// TIA Portal project "exografcet2" (V16)

(* hardware
DEVICE "Station S7-1200_1"  S7-1200 Station
   slot 0: "Châssis_0"  S7-1200 Rack  Rack  V1.0
   slot 1: "PLC_1"  CPU 1214C AC/DC/Rly  6ES7 214-1BG40-0XB0  V4.4
*)

// ===== PLC "PLC_1"  CPU 1214C AC/DC/Rly =====

VAR_GLOBAL   // PLC tag table "Table de variables standard"
   "MARCHE" AT %I0.0 : Bool;
   "ARRET" AT %I0.1 : Bool;
   "moteur" AT %Q0.0 : Bool;
   "H1" AT %Q0.1 : Bool;
   "H2" AT %Q0.2 : Bool;
END_VAR

ORGANIZATION_BLOCK "Main"   // OB1, LAD, ProgramCycle
TITLE = "Main Program Sweep (Cycle)"
{ S7_Optimized_Access := 'TRUE' }
VERSION : 0.1
   VAR_INPUT
      Initial_Call : Bool;   // Initial call of this OB
      Remanence : Bool;   // =True, if remanent data are available
   END_VAR
BEGIN

REGION Network 1
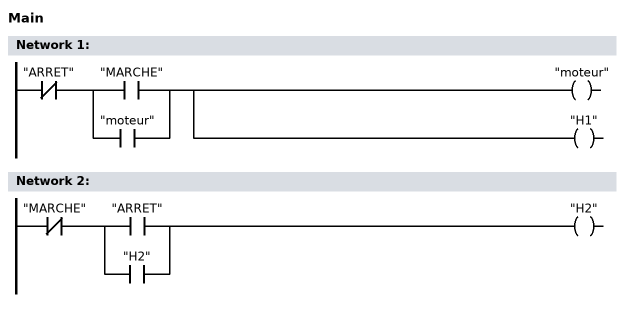
   RUNG wire#powerrail
      I_Contact( "ARRET" )
      wire#w1
      Contact( "MARCHE" )
      wire#w2
      Coil( "moteur" )
   END_RUNG
   RUNG wire#w1
      Contact( "moteur" )
   END_RUNG wire#w2
   RUNG wire#w2
      Coil( "H1" )
   END_RUNG
   // the same network as SCL:
   "moteur" := NOT "ARRET" AND ("MARCHE" OR "moteur");
   "H1" := "moteur";
END_REGION

REGION Network 2
   RUNG wire#powerrail
      I_Contact( "MARCHE" )
      wire#w1
      Contact( "ARRET" )
      wire#w2
      Coil( "H2" )
   END_RUNG
   RUNG wire#w1
      Contact( "H2" )
   END_RUNG wire#w2
   // the same network as SCL:
   "H2" := NOT "MARCHE" AND ("ARRET" OR "H2");
END_REGION
END_ORGANIZATION_BLOCK